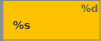
VISUALIZATION FRM_SafetyElement  // 101x41
VAR_INPUT
   nIndex: USINT;
   nOffset: USINT;
END_VAR
    Rectangle (3,0 98x41)
    Textfield (10,10 91x31), "%s", text variable: Motion_Safety.stSafety.stOut.astDiagnosticElement[nIndex + nOffset].sName
    Rectangle (0,0 3x41), colour toggle: Motion_Safety.fbMotionSafety.stPNOZEtherCATDiagIn.astDiagnosticElementsIn[nIndex + nOffset].nLow.b1
    Textfield (80,3 21x11), "%d", text variable: nIndex + nOffset
    Rectangle (0,0 3x41), invisible if: Motion_Safety.fbMotionSafety.stPNOZEtherCATDiagIn.astDiagnosticElementsIn[nIndex + nOffset].nLow.b0
    Rectangle (0,0 101x41)
        OnMouseUp: execute { GVL_Safety.nHMIDiagWordIndex := nIndex + nOffset; }
        OnMouseUp: OpenDialog Dialog=FRM_WordDiagnostic, OpenModal=True, OpenCentered=True
END_VISUALIZATION

(* stored: Version 1.1.0.1
   Visu FRM_SafetyElement: Id {b603ab46-f5d8-02c5-2b4b-4ca604f5117d} *)
